(* LS Electric XG5000 project: ROUND *)
(* PLC LSPLC *)

PROGRAM NewProgram (* task: 스캔 프로그램 *)
VAR
    BothCounter : CTUD_DINT;
    DownCounter : CTD_DINT;
    Fall : F_TRIG;
    FF : FF;
    OffTimer : TOF;
    OnTimer : TON;
    PulseTimer : TP;
    ResetLatch : RS;
    Rise : R_TRIG;
    SetLatch : SR;
    UpCounter : CTU_DINT;
END_VAR
VAR
    _t1 : BOOL;
END_VAR

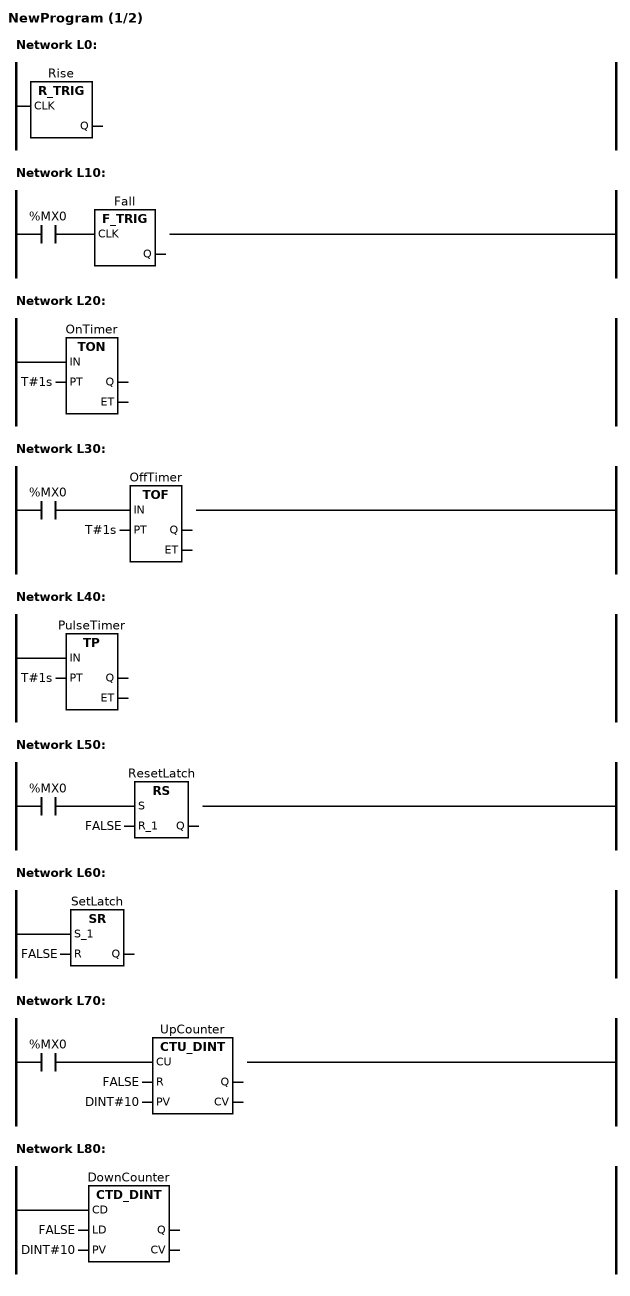
(* Rung L0 *)
Rise(CLK := TRUE);
(* Rung L10 *)
Fall(CLK := %MX0);
(* Rung L20 *)
OnTimer(IN := TRUE, PT := T#1s);
(* Rung L30 *)
OffTimer(IN := %MX0, PT := T#1s);
(* Rung L40 *)
PulseTimer(IN := TRUE, PT := T#1s);
(* Rung L50 *)
ResetLatch(S := %MX0, R_1 := FALSE);
(* Rung L60 *)
SetLatch(S_1 := TRUE, R := FALSE);
(* Rung L70 *)
UpCounter(CU := %MX0, R := FALSE, PV := DINT#10);
(* Rung L80 *)
DownCounter(CD := TRUE, LD := FALSE, PV := DINT#10);

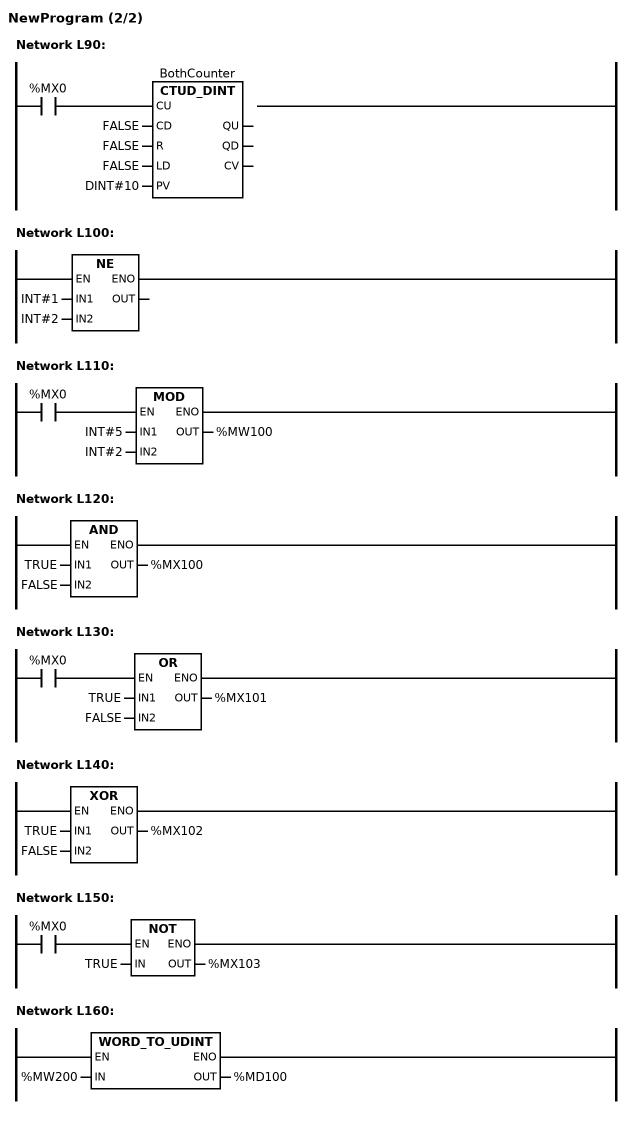
(* Rung L90 *)
BothCounter(CU := %MX0, CD := FALSE, R := FALSE, LD := FALSE, PV := DINT#10);
(* Rung L100 *)
_t1 := INT#1 <> INT#2;
(* Rung L110 *)
IF %MX0 THEN %MW100 := INT#5 MOD INT#2; END_IF;
(* Rung L120 *)
%MX100 := TRUE AND FALSE;
(* Rung L130 *)
IF %MX0 THEN %MX101 := TRUE OR FALSE; END_IF;
(* Rung L140 *)
%MX102 := TRUE XOR FALSE;
(* Rung L150 *)
IF %MX0 THEN %MX103 := NOT TRUE; END_IF;
(* Rung L160 *)
%MD100 := WORD_TO_UDINT(%MW200);
END_PROGRAM